{region 'Documentation'}
(*!
<summary>Check that the token count is outside the inclusive Minimum..Maximum range.</summary>
<description>

StartIndex is an absolute declared IN index, not an offset. Length selects 1..255
elements; the complete selected range must fit IN. Invalid references or ranges report
Error.

Keep supplied arrays stable for the call. Input data is read, not copied or retained as a
snapshot.

Counts the currently selected region on evaluation, not occurrences across cycles.
TokenCount exposes the last computed count. Inclusive range bounds must be ordered; reversed
bounds report Error.

Token is the complete nonempty array pattern starting at its own lower bound and must fit
the selected search range; otherwise Error. Array token matching is exact.

Matches do not overlap: searching resumes after the whole matched token.

</description>
*)
{endregion}
FUNCTION_BLOCK AssertArrayTokenCntNotInRange_Byte EXTENDS AssertionBase
VAR_INPUT
    StartIndex : DINT; //! First selected index in IN; uses the array's declared index range, not a zero-based offset.
    Length : USINT; //! Number of selected elements starting at StartIndex; must fit the array range; valid range 1..255.
    Minimum : UINT; //! Inclusive lower bound of the comparison; for a range, must not exceed Maximum.
    Maximum : UINT; //! Inclusive upper bound of the comparison; for a range, must not be below Minimum.
END_VAR
VAR_IN_OUT CONSTANT
    IN : ARRAY[*] OF BYTE; //! Keep the searched data stable during the call.
    Token : ARRAY[*] OF BYTE; //! Read-only nonempty token; keep stable during the call and within the selected search length.
END_VAR
VAR
    FTokenCount : UINT;
END_VAR

SUPER^();

{region 'Documentation'}
(*!
<summary>Validate configuration, count tokens and apply the count predicate.</summary>
*)
{endregion}
METHOD PROTECTED Assert
VAR
    InLowerIndex : DINT;
    InUpperIndex : DINT;
    EndIndex : LINT;
    TokenLowerIndex : DINT;
    TokenUpperIndex : DINT;
    TokenLength : LINT;
    Message : STRING(GVL_Constants.MessageLength);
END_VAR
IF NOT EvaluationActive THEN
    RETURN;
END_IF;

IF Result = E_Result.Error THEN
    RETURN;
END_IF;

// C0371: FB input is checked before any reference access.
{warning disable C0371}
IF NOT __ISVALIDREF(IN) THEN
    FTokenCount := 0;
    Error(Message := 'Assertion error: IN reference is invalid.');
    RETURN;
END_IF;

IF NOT __ISVALIDREF(Token) THEN
    FTokenCount := 0;
    Error(Message := 'Assertion error: Token reference is invalid.');
    RETURN;
END_IF;

TokenLowerIndex := LOWER_BOUND(Token, 1);
TokenUpperIndex := UPPER_BOUND(Token, 1);
TokenLength := DINT_TO_LINT(TokenUpperIndex) - DINT_TO_LINT(TokenLowerIndex) + 1;
IF (TokenLength <= 0) OR (TokenLength > USINT_TO_LINT(Length)) THEN
    FTokenCount := 0;
    Message := CONCAT('Assertion error: invalid token length. TokenLength = ',
        LINT_TO_STRING(TokenLength));
    Message := CONCAT(Message, ', Length = ');
    Message := CONCAT(Message, USINT_TO_STRING(Length));
    Error(Message := Message);
    RETURN;
END_IF;

InLowerIndex := LOWER_BOUND(IN, 1);
InUpperIndex := UPPER_BOUND(IN, 1);
EndIndex := DINT_TO_LINT(StartIndex) + USINT_TO_LINT(Length) - 1;
IF (Length = 0)
    OR (StartIndex < InLowerIndex) OR (StartIndex > InUpperIndex)
    OR (EndIndex > DINT_TO_LINT(InUpperIndex)) THEN
    FTokenCount := 0;
    Message := CONCAT('Assertion error: invalid search range. StartIndex = ',
        DINT_TO_STRING(StartIndex));
    Message := CONCAT(Message, ', Length = ');
    Message := CONCAT(Message, USINT_TO_STRING(Length));
    Error(Message := Message);
    RETURN;
END_IF;

IF Minimum > Maximum THEN
    FTokenCount := 0;
    Message := CONCAT('Assertion error: reversed token count bounds. Minimum = ',
        UINT_TO_STRING(Minimum));
    Message := CONCAT(Message, ', Maximum = ');
    Message := CONCAT(Message, UINT_TO_STRING(Maximum));
    Error(Message := Message);
    RETURN;
END_IF;

IF Result = E_Result.Failed THEN
    RETURN;
END_IF;

FTokenCount := CountArrayTokens_Byte(StartIndex := StartIndex,
    Length := Length,
    Token := Token,
    IN := IN);

IF (FTokenCount >= Minimum) AND (FTokenCount <= Maximum) THEN
    Message := CONCAT('Assertion failed: array token count violates NotInRange. Actual = ',
        UINT_TO_STRING(FTokenCount));
    Message := CONCAT(Message, ', Minimum = ');
    Message := CONCAT(Message, UINT_TO_STRING(Minimum));
    Message := CONCAT(Message, ', Maximum = ');
    Message := CONCAT(Message, UINT_TO_STRING(Maximum));
    Message := CONCAT(Message, ', TokenRange = [');
    Message := CONCAT(Message, DINT_TO_STRING(TokenLowerIndex));
    Message := CONCAT(Message, '..');
    Message := CONCAT(Message, DINT_TO_STRING(TokenUpperIndex));
    Message := CONCAT(Message, ']');
    Fail(Message := Message);
    RETURN;
END_IF;

Pass();
{warning restore C0371}
END_METHOD

{region 'Documentation'}
(*!
<summary>Clear the retained count on framework reset.</summary>
*)
{endregion}
METHOD PROTECTED ResetAssertion
FTokenCount := 0;
END_METHOD

{region 'Documentation'}
(*!
<summary>Return the most recently evaluated token count.</summary>
<description>

Counts occurrences in one selected array region, not across PLC cycles. Retained while
disabled or after Failed; reset and detected configuration errors clear it. Reading this
property does not search the array.

</description>
*)
{endregion}
{attribute 'monitoring' := 'call'}
PROPERTY PUBLIC TokenCount : UINT //! Return the most recently evaluated token count.
GET // PUBLIC
TokenCount := FTokenCount;
END_GET
END_PROPERTY

END_FUNCTION_BLOCK

(* stored: Version 1.1.0.1
   POU AssertArrayTokenCntNotInRange_Byte: Id {941df28f-4e9b-43b3-8c98-c5fc275445af}, SpecialFunc None
   Folder Internal: Id {443d7111-6fe5-4621-95af-b7d028a38063}
   Method Assert: Id {31a692ab-36df-4d12-83cc-3160537c78c4}
   Method ResetAssertion: Id {f746e717-eb41-48a7-801d-ea283c46790a}
   Property TokenCount: Id {3ec77a77-9bc3-4865-b786-3bec3027bb50}
   Get Get: Id {1e83eba4-1046-4dec-82f5-7cad4ad0b6ad} *)
